// TIA Portal V19 export
// export: Created 2026-10-15T10:10:17.0177146Z, ExportSetting WithDefaults, DisplayName Totally Integrated Automation Portal, DisplayVersion V19, DisplayName TIA Portal Openness, DisplayVersion V19, DisplayName TIA Portal Version Control Interface, DisplayVersion V19, DisplayName STEP 7 Professional, DisplayVersion V19, DisplayName STEP 7 Safety, DisplayVersion V19, DisplayName WinCC Basic/Comfort/Advanced, DisplayVersion V19, DisplayName WinCC Unified, DisplayVersion V19
DATA_BLOCK "ROLL_DB15"   // DB4
{ S7_Optimized_Access := 'TRUE' }
VERSION : 0.1
// stored: AutoNumber true, DBAccessibleFromOPCUA true, DBAccessibleFromWebserver true, IsOnlyStoredInLoadMemory false, IsRetainMemResEnabled false, IsWriteProtectedInAS false, MemoryReserve 100
   VAR
      DW : Array[0..131] of Word;
   END_VAR
BEGIN
   DW[0..16] := WORD#16#FFFF;
   DW[17] := WORD#16#3360;
   DW[18..23] := WORD#16#FFFF;
   DW[24] := WORD#16#1010;
   DW[25] := WORD#16#1020;
   DW[26..30] := WORD#16#FFFF;
   DW[31..32] := WORD#16#3120;
   DW[33] := WORD#16#2900;
   DW[34..52] := WORD#16#FFFF;
   DW[53..54] := WORD#16#2120;
   DW[55] := WORD#16#1010;
   DW[56] := WORD#16#2060;
   DW[57] := WORD#16#FFFF;
   DW[58..59] := WORD#16#3180;
   DW[60] := WORD#16#2060;
   DW[61..62] := WORD#16#2600;
   DW[63] := WORD#16#2010;
   DW[64] := WORD#16#FFFF;
   DW[65] := WORD#16#2015;
   DW[66] := WORD#16#FFFF;
   DW[67] := WORD#16#1050;
   DW[68..74] := WORD#16#FFFF;
   DW[75] := WORD#16#2600;
   DW[76] := WORD#16#FFFF;
   DW[77] := WORD#16#2300;
   DW[78..84] := WORD#16#FFFF;
   DW[85] := WORD#16#2120;
   DW[86..101] := WORD#16#FFFF;
   DW[102..103] := WORD#16#2300;
   DW[104..105] := WORD#16#FFFF;
   DW[106] := WORD#16#2010;
   DW[107] := WORD#16#2015;
   DW[108..114] := WORD#16#FFFF;
   DW[115..117] := WORD#16#1050;
   DW[118..126] := WORD#16#FFFF;
   DW[127] := WORD#16#0038;
   DW[128..129] := WORD#16#0011;
   DW[130] := WORD#16#3360;
END_DATA_BLOCK
